// TIA Portal project "S7-1200-Single-Pump-Station" (V17)

(* hardware
DEVICE "S7-1200 station_1"  S7-1200 Station
   slot 0: "Rack_0"  S7-1200 Rack  Rack  V1.0
   slot 1: "PLC_1"  CPU 1212C DC/DC/DC  6ES7 212-1AE40-0XB0  V4.2
DEVICE "HMI_1"  TP700 Comfort
   slot 0: "HMI_1"  TP700 Comfort  6AV2 124-0GC01-0AX0  17.0.0.0
   slot 1: "HMI_RT_1"  TP700 Comfort  6AV2 124-0GC01-0AX0  17.0.0.0
   slot 5: "HMI_1.IE_CP_1"  PROFINET Interface  17.0.0.0
      slot 1: "PROFINET Interface_1"  PROFINET Interface
         slot 1: "Port_1"  Port
         slot 2: "Port_2"  Port
   slot 7: "HMI_1.MPI/DP_CP_1"  MPI/DP Interface  17.0.0.0
*)

// ===== PLC "PLC_1"  CPU 1212C DC/DC/DC =====

VAR_GLOBAL   // PLC tag table "Default tag table"
   "Clock_Byte" AT %MB100 : Byte;
   "Clock_10Hz" AT %M100.0 : Bool;
   "Clock_5Hz" AT %M100.1 : Bool;
   "Clock_2.5Hz" AT %M100.2 : Bool;
   "Clock_2Hz" AT %M100.3 : Bool;
   "Clock_1.25Hz" AT %M100.4 : Bool;
   "Clock_1Hz" AT %M100.5 : Bool;
   "Clock_0.625Hz" AT %M100.6 : Bool;
   "Clock_0.5Hz" AT %M100.7 : Bool;
   "AL" AT %I0.5 : Bool;
   "LSL" AT %I0.3 : Bool;
   "LSH" AT %I0.4 : Bool;
   "S1Auto" AT %I0.0 : Bool;
   "S2" AT %I0.2 : Bool;
   "LT" AT %IW64 : Int;
   "L1" AT %Q0.0 : Bool;
   "L2" AT %Q0.1 : Bool;
   "P1" AT %Q0.2 : Bool;
   "S1Hand" AT %I0.1 : Bool;
END_VAR

DATA_BLOCK "Random Generator DB"   // DB1
{ S7_Optimized_Access := 'TRUE' }
VERSION : 0.1
// stored: InstanceOfName Random Inflow Generator
"Random Inflow Generator"
BEGIN
END_DATA_BLOCK

DATA_BLOCK "Well DB"   // DB3
{ S7_Optimized_Access := 'TRUE' }
VERSION : 0.1
// stored: InstanceOfName Well Simulation
"Well Simulation"
BEGIN
END_DATA_BLOCK

DATA_BLOCK "Main DB"   // DB4
{ S7_Optimized_Access := 'TRUE' }
VERSION : 0.1
   VAR
      RandomInflow : Real;
      ActualInflow : Real;
      ActualOutflow : Real;
      S1AutoHMI : Bool;
      S1HandHMI : Bool;
      S2HMI : Bool;
      AutoMode : Bool;
      HandMode : Bool;
      ServiceMode : Bool;
      LevelPercent : Real;
      HighLevelReached : Bool;
      AutoPumpLatch : Bool;
      LSHHMI : Bool;
      LSLHMI : Bool;
      AlarmMode : Bool;
      HighLevelSetpoint : Real := 50.0;
      LowLevelSetpoint : Real := 20.0;
      ResetSetpoints : Bool;
      AlarmHelp : Bool := false;
      LTMeters : Real;
      ALHMI : Bool;
      PumpFault : Bool;
      HMIAlarmWord : Word;
      HighSetpointPrevious : Real := 50.0;
      LowSetpointPrevious : Real := 20.0;
      LTNormalized : Real;
      LTAnalogPercent : Real;
      SimulationMode : Bool;
      PumpStartRequest : Bool;
      PumpSafety : Bool;
      LevelInLiters : Real;
   END_VAR
BEGIN
END_DATA_BLOCK

// folder: System blocks/Program resources

DATA_BLOCK "IEC_Timer_0_DB"   // DB2
{ S7_Optimized_Access := 'TRUE' }
AUTHOR : Simatic
FAMILY : IEC
NAME : IEC_TMR
VERSION : 1.0
// stored: InstanceOfName IEC_TIMER
"IEC_TIMER"
BEGIN
END_DATA_BLOCK

DATA_BLOCK "IEC_Timer_0_DB_2"   // DB6
{ S7_Optimized_Access := 'TRUE' }
AUTHOR : Simatic
FAMILY : IEC
NAME : IEC_TMR
VERSION : 1.0
// stored: InstanceOfName IEC_TIMER
"IEC_TIMER"
BEGIN
END_DATA_BLOCK

// folder: (top level)

FUNCTION_BLOCK "Random Inflow Generator"   // FB1, LAD
{ S7_Optimized_Access := 'TRUE' }
VERSION : 0.1
   VAR_OUTPUT
      RandomInflow : Real;
   END_VAR
   VAR
      TimeStatus : Int;
      SystemTime : DTL;
      RandomValue : Int;
   END_VAR
BEGIN

REGION Network 1: System Time Acquisition
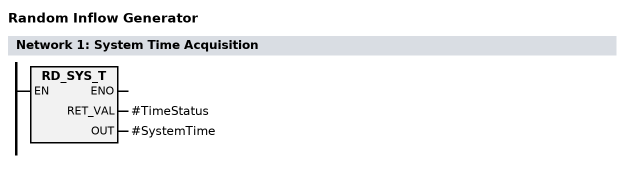
   #TimeStatus := RD_SYS_T(OUT => #SystemTime);
END_REGION

REGION Network 2 (SCL): Random Value Generation
   IF #TimeStatus = 0 THEN
       #RandomValue :=
       UDINT_TO_INT(
                     #SystemTime.NANOSECOND MOD UDINT#3
       ) + 1;
   END_IF;
END_REGION

REGION Network 3 (SCL): Random Inflow Rate Selection
   IF #RandomValue = 1 THEN
       #RandomInflow := 10.0;
   ELSIF #RandomValue = 2 THEN
       #RandomInflow := 15.0;
   ELSE
       #RandomInflow := 7.0;
   END_IF;
END_REGION
END_FUNCTION_BLOCK

FUNCTION_BLOCK "Well Simulation"   // FB2, SCL
{ S7_Optimized_Access := 'TRUE' }
VERSION : 0.1
   VAR_INPUT
      CycleTime : Real := 0.1;
      Inflow : Real;
      Outflow : Real;
   END_VAR
   VAR
      TankLevel : Real;
      ActualInflow : Real;
      ActualOutflow : Real;
      "TankLevel%" : Real;
   END_VAR
BEGIN
   #ActualOutflow := #Outflow * #CycleTime;
   #ActualInflow := #Inflow * #CycleTime;

   #TankLevel := #TankLevel + (#ActualInflow - #ActualOutflow);

   IF #TankLevel > 1250.0 THEN
       #TankLevel := 1250.0;
   END_IF;

   IF #TankLevel < 0.0 THEN
       #TankLevel := 0.0;
   END_IF;

   #"TankLevel%" := (#TankLevel / 1250.0) * 100.0;
END_FUNCTION_BLOCK

ORGANIZATION_BLOCK "Main"   // OB1, LAD, ProgramCycle
TITLE = "Main Program Sweep (Cycle)"
{ S7_Optimized_Access := 'TRUE' }
VERSION : 0.1
   VAR_INPUT
      Initial_Call : Bool;   // Initial call of this OB
      Remanence : Bool;   // =True, if remanent data are available
   END_VAR
BEGIN

REGION Network 1: LT Analog Input Scaling
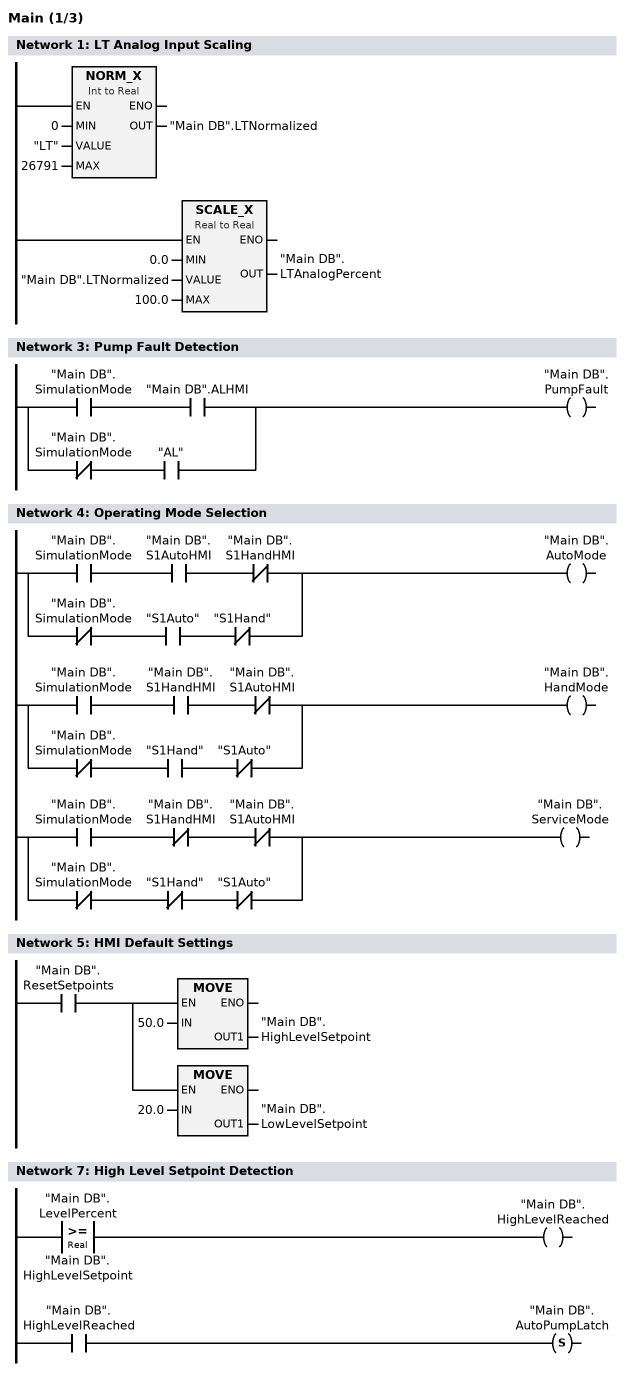
   RUNG wire#powerrail
      { S7_Templates := "[SrcType := Int, DestType := Real]" } Normalize(min := 0, value := "LT", max := 26791, out => "Main DB".LTNormalized)
   END_RUNG
   RUNG wire#powerrail
      { S7_Templates := "[SrcType := Real, DestType := Real]" } Scale(min := 0.0, value := "Main DB".LTNormalized, max := 100.0, out => "Main DB".LTAnalogPercent)
   END_RUNG
   // the same network as SCL:
   "Main DB".LTNormalized := NORM_X(MIN := 0, VALUE := "LT", MAX := 26791);
   "Main DB".LTAnalogPercent := SCALE_X(MIN := 0.0, VALUE := "Main DB".LTNormalized, MAX := 100.0);
END_REGION

REGION Network 2 (SCL): LT Source Selection and Level Conversion
   IF "Main DB".SimulationMode THEN
       "Main DB".LevelPercent := "Well DB"."TankLevel%";
       "Main DB".LevelInLiters := "Well DB".TankLevel;
   ELSE
       "Main DB".LevelPercent := "Main DB".LTAnalogPercent;
       "Main DB".LevelInLiters := ("Main DB".LevelPercent / 100.0) * 1250.0;
   END_IF;

   "Main DB".LTMeters := ("Main DB".LevelPercent * 2.5) / 100.0;
END_REGION

REGION Network 3: Pump Fault Detection
   RUNG wire#powerrail
      Contact( "Main DB".SimulationMode )
      Contact( "Main DB".ALHMI )
      wire#w1
      Coil( "Main DB".PumpFault )
   END_RUNG
   RUNG wire#powerrail
      I_Contact( "Main DB".SimulationMode )
      Contact( "AL" )
   END_RUNG wire#w1
   // the same network as SCL:
   "Main DB".PumpFault := ("Main DB".SimulationMode AND "Main DB".ALHMI) OR (NOT "Main DB".SimulationMode AND "AL");
END_REGION

REGION Network 4: Operating Mode Selection
   RUNG wire#powerrail
      Contact( "Main DB".SimulationMode )
      Contact( "Main DB".S1AutoHMI )
      I_Contact( "Main DB".S1HandHMI )
      wire#w1
      Coil( "Main DB".AutoMode )
   END_RUNG
   RUNG wire#powerrail
      I_Contact( "Main DB".SimulationMode )
      Contact( "S1Auto" )
      I_Contact( "S1Hand" )
   END_RUNG wire#w1
   RUNG wire#powerrail
      Contact( "Main DB".SimulationMode )
      Contact( "Main DB".S1HandHMI )
      I_Contact( "Main DB".S1AutoHMI )
      wire#w2
      Coil( "Main DB".HandMode )
   END_RUNG
   RUNG wire#powerrail
      I_Contact( "Main DB".SimulationMode )
      Contact( "S1Hand" )
      I_Contact( "S1Auto" )
   END_RUNG wire#w2
   RUNG wire#powerrail
      Contact( "Main DB".SimulationMode )
      I_Contact( "Main DB".S1HandHMI )
      I_Contact( "Main DB".S1AutoHMI )
      wire#w3
      Coil( "Main DB".ServiceMode )
   END_RUNG
   RUNG wire#powerrail
      I_Contact( "Main DB".SimulationMode )
      I_Contact( "S1Hand" )
      I_Contact( "S1Auto" )
   END_RUNG wire#w3
   // the same network as SCL:
   "Main DB".AutoMode := ("Main DB".SimulationMode AND "Main DB".S1AutoHMI AND NOT "Main DB".S1HandHMI) OR (NOT "Main DB".SimulationMode AND "S1Auto" AND NOT "S1Hand");
   "Main DB".HandMode := ("Main DB".SimulationMode AND "Main DB".S1HandHMI AND NOT "Main DB".S1AutoHMI) OR (NOT "Main DB".SimulationMode AND "S1Hand" AND NOT "S1Auto");
   "Main DB".ServiceMode := ("Main DB".SimulationMode AND NOT "Main DB".S1HandHMI AND NOT "Main DB".S1AutoHMI) OR (NOT "Main DB".SimulationMode AND NOT "S1Hand" AND NOT "S1Auto");
END_REGION

REGION Network 5: HMI Default Settings
   RUNG wire#powerrail
      Contact( "Main DB".ResetSetpoints )
      wire#w1
      Move(in := 50.0, out1 => "Main DB".HighLevelSetpoint)
   END_RUNG
   RUNG wire#w1
      Move(in := 20.0, out1 => "Main DB".LowLevelSetpoint)
   END_RUNG
   // the same network as SCL:
   IF "Main DB".ResetSetpoints THEN
       "Main DB".HighLevelSetpoint := 50.0;
       "Main DB".LowLevelSetpoint := 20.0;
   END_IF;
END_REGION

REGION Network 6 (SCL): HMI Setpoint Validation

   IF "Main DB".LowLevelSetpoint <> "Main DB".LowSetpointPrevious THEN

       "Main DB".LowLevelSetpoint := LIMIT(
                                           MN := 0.0,
                                           IN := "Main DB".LowLevelSetpoint,
                                           MX := "Main DB".HighLevelSetpoint - 5.0
       );

   ELSIF "Main DB".HighLevelSetpoint <> "Main DB".HighSetpointPrevious THEN

       "Main DB".HighLevelSetpoint := LIMIT(
                                            MN := "Main DB".LowLevelSetpoint + 5.0,
                                            IN := "Main DB".HighLevelSetpoint,
                                            MX := 100.0
       );

   END_IF;

   "Main DB".HighSetpointPrevious := "Main DB".HighLevelSetpoint;
   "Main DB".LowSetpointPrevious := "Main DB".LowLevelSetpoint;
END_REGION

REGION Network 7: High Level Setpoint Detection
   RUNG wire#powerrail
      { S7_Templates := "SrcType := Real" } GE_Contact(in1 := "Main DB".LevelPercent, in2 := "Main DB".HighLevelSetpoint)
      Coil( "Main DB".HighLevelReached )
   END_RUNG
   RUNG wire#powerrail
      Contact( "Main DB".HighLevelReached )
      S_Coil( "Main DB".AutoPumpLatch )
   END_RUNG
   // the same network as SCL:
   "Main DB".HighLevelReached := "Main DB".LevelPercent >= "Main DB".HighLevelSetpoint;
   IF "Main DB".HighLevelReached THEN "Main DB".AutoPumpLatch := TRUE; END_IF;
END_REGION

REGION Network 8: Low Level Setpoint Reset
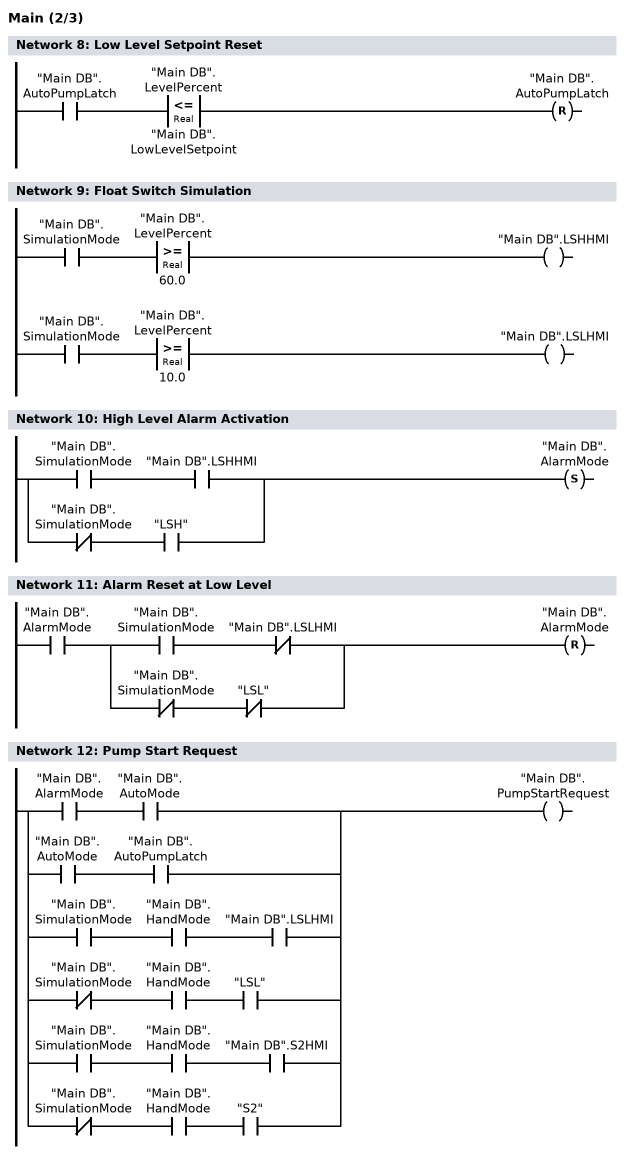
   RUNG wire#powerrail
      Contact( "Main DB".AutoPumpLatch )
      { S7_Templates := "SrcType := Real" } LE_Contact(in1 := "Main DB".LevelPercent, in2 := "Main DB".LowLevelSetpoint)
      R_Coil( "Main DB".AutoPumpLatch )
   END_RUNG
   // the same network as SCL:
   IF "Main DB".AutoPumpLatch AND ("Main DB".LevelPercent <= "Main DB".LowLevelSetpoint) THEN
       "Main DB".AutoPumpLatch := FALSE;
   END_IF;
END_REGION

REGION Network 9: Float Switch Simulation
   RUNG wire#powerrail
      Contact( "Main DB".SimulationMode )
      { S7_Templates := "SrcType := Real" } GE_Contact(in1 := "Main DB".LevelPercent, in2 := 60.0)
      Coil( "Main DB".LSHHMI )
   END_RUNG
   RUNG wire#powerrail
      Contact( "Main DB".SimulationMode )
      { S7_Templates := "SrcType := Real" } GE_Contact(in1 := "Main DB".LevelPercent, in2 := 10.0)
      Coil( "Main DB".LSLHMI )
   END_RUNG
   // the same network as SCL:
   "Main DB".LSHHMI := "Main DB".SimulationMode AND ("Main DB".LevelPercent >= 60.0);
   "Main DB".LSLHMI := "Main DB".SimulationMode AND ("Main DB".LevelPercent >= 10.0);
END_REGION

REGION Network 10: High Level Alarm Activation
   RUNG wire#powerrail
      Contact( "Main DB".SimulationMode )
      Contact( "Main DB".LSHHMI )
      wire#w1
      S_Coil( "Main DB".AlarmMode )
   END_RUNG
   RUNG wire#powerrail
      I_Contact( "Main DB".SimulationMode )
      Contact( "LSH" )
   END_RUNG wire#w1
   // the same network as SCL:
   IF ("Main DB".SimulationMode AND "Main DB".LSHHMI) OR (NOT "Main DB".SimulationMode AND "LSH") THEN
       "Main DB".AlarmMode := TRUE;
   END_IF;
END_REGION

REGION Network 11: Alarm Reset at Low Level
   RUNG wire#powerrail
      Contact( "Main DB".AlarmMode )
      wire#w1
      Contact( "Main DB".SimulationMode )
      I_Contact( "Main DB".LSLHMI )
      wire#w2
      R_Coil( "Main DB".AlarmMode )
   END_RUNG
   RUNG wire#w1
      I_Contact( "Main DB".SimulationMode )
      I_Contact( "LSL" )
   END_RUNG wire#w2
   // the same network as SCL:
   IF "Main DB".AlarmMode AND (("Main DB".SimulationMode AND NOT "Main DB".LSLHMI) OR (NOT "Main DB".SimulationMode AND NOT "LSL")) THEN
       "Main DB".AlarmMode := FALSE;
   END_IF;
END_REGION

REGION Network 12: Pump Start Request
   RUNG wire#powerrail
      Contact( "Main DB".AlarmMode )
      Contact( "Main DB".AutoMode )
      wire#w1
      Coil( "Main DB".PumpStartRequest )
   END_RUNG
   RUNG wire#powerrail
      Contact( "Main DB".AutoMode )
      Contact( "Main DB".AutoPumpLatch )
   END_RUNG wire#w1
   RUNG wire#powerrail
      Contact( "Main DB".SimulationMode )
      Contact( "Main DB".HandMode )
      Contact( "Main DB".LSLHMI )
   END_RUNG wire#w1
   RUNG wire#powerrail
      I_Contact( "Main DB".SimulationMode )
      Contact( "Main DB".HandMode )
      Contact( "LSL" )
   END_RUNG wire#w1
   RUNG wire#powerrail
      Contact( "Main DB".SimulationMode )
      Contact( "Main DB".HandMode )
      Contact( "Main DB".S2HMI )
   END_RUNG wire#w1
   RUNG wire#powerrail
      I_Contact( "Main DB".SimulationMode )
      Contact( "Main DB".HandMode )
      Contact( "S2" )
   END_RUNG wire#w1
   // the same network as SCL:
   "Main DB".PumpStartRequest := ("Main DB".AlarmMode AND "Main DB".AutoMode) OR ("Main DB".AutoMode AND "Main DB".AutoPumpLatch) OR ("Main DB".SimulationMode AND "Main DB".HandMode AND "Main DB".LSLHMI) OR (NOT "Main DB".SimulationMode AND "Main DB".HandMode AND "LSL") OR ("Main DB".SimulationMode AND "Main DB".HandMode AND "Main DB".S2HMI) OR (NOT "Main DB".SimulationMode AND "Main DB".HandMode AND "S2");
END_REGION

REGION Network 13: Pump Safety Interlocks
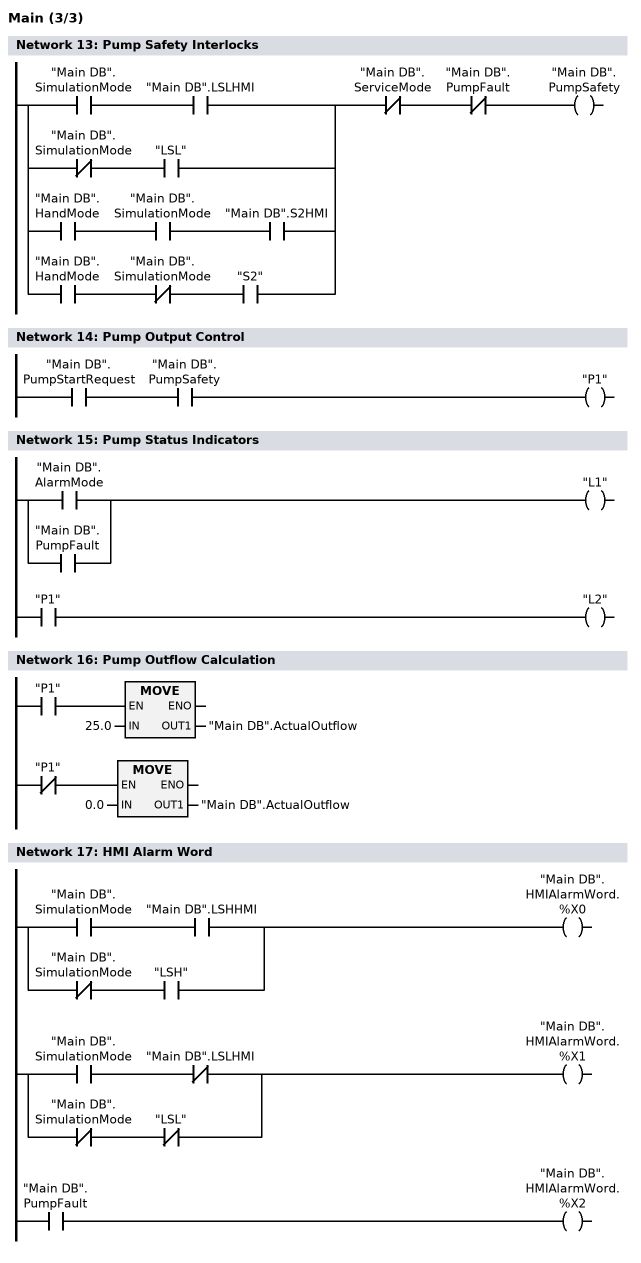
   RUNG wire#powerrail
      Contact( "Main DB".SimulationMode )
      Contact( "Main DB".LSLHMI )
      wire#w1
      I_Contact( "Main DB".ServiceMode )
      I_Contact( "Main DB".PumpFault )
      Coil( "Main DB".PumpSafety )
   END_RUNG
   RUNG wire#powerrail
      I_Contact( "Main DB".SimulationMode )
      Contact( "LSL" )
   END_RUNG wire#w1
   RUNG wire#powerrail
      Contact( "Main DB".HandMode )
      Contact( "Main DB".SimulationMode )
      Contact( "Main DB".S2HMI )
   END_RUNG wire#w1
   RUNG wire#powerrail
      Contact( "Main DB".HandMode )
      I_Contact( "Main DB".SimulationMode )
      Contact( "S2" )
   END_RUNG wire#w1
   // the same network as SCL:
   "Main DB".PumpSafety := (("Main DB".SimulationMode AND "Main DB".LSLHMI) OR (NOT "Main DB".SimulationMode AND "LSL") OR ("Main DB".HandMode AND "Main DB".SimulationMode AND "Main DB".S2HMI) OR ("Main DB".HandMode AND NOT "Main DB".SimulationMode AND "S2")) AND NOT "Main DB".ServiceMode AND NOT "Main DB".PumpFault;
END_REGION

REGION Network 14: Pump Output Control
   RUNG wire#powerrail
      Contact( "Main DB".PumpStartRequest )
      Contact( "Main DB".PumpSafety )
      Coil( "P1" )
   END_RUNG
   // the same network as SCL:
   "P1" := "Main DB".PumpStartRequest AND "Main DB".PumpSafety;
END_REGION

REGION Network 15: Pump Status Indicators
   RUNG wire#powerrail
      Contact( "Main DB".AlarmMode )
      wire#w1
      Coil( "L1" )
   END_RUNG
   RUNG wire#powerrail
      Contact( "Main DB".PumpFault )
   END_RUNG wire#w1
   RUNG wire#powerrail
      Contact( "P1" )
      Coil( "L2" )
   END_RUNG
   // the same network as SCL:
   "L1" := "Main DB".AlarmMode OR "Main DB".PumpFault;
   "L2" := "P1";
END_REGION

REGION Network 16: Pump Outflow Calculation
   RUNG wire#powerrail
      Contact( "P1" )
      Move(in := 25.0, out1 => "Main DB".ActualOutflow)
   END_RUNG
   RUNG wire#powerrail
      I_Contact( "P1" )
      Move(in := 0.0, out1 => "Main DB".ActualOutflow)
   END_RUNG
   // the same network as SCL:
   IF "P1" THEN "Main DB".ActualOutflow := 25.0; END_IF;
   IF NOT "P1" THEN "Main DB".ActualOutflow := 0.0; END_IF;
END_REGION

REGION Network 17: HMI Alarm Word
   RUNG wire#powerrail
      Contact( "Main DB".SimulationMode )
      Contact( "Main DB".LSHHMI )
      wire#w1
      Coil( "Main DB".HMIAlarmWord.%X0 )
   END_RUNG
   RUNG wire#powerrail
      I_Contact( "Main DB".SimulationMode )
      Contact( "LSH" )
   END_RUNG wire#w1
   RUNG wire#powerrail
      Contact( "Main DB".SimulationMode )
      I_Contact( "Main DB".LSLHMI )
      wire#w2
      Coil( "Main DB".HMIAlarmWord.%X1 )
   END_RUNG
   RUNG wire#powerrail
      I_Contact( "Main DB".SimulationMode )
      I_Contact( "LSL" )
   END_RUNG wire#w2
   RUNG wire#powerrail
      Contact( "Main DB".PumpFault )
      Coil( "Main DB".HMIAlarmWord.%X2 )
   END_RUNG
   // the same network as SCL:
   "Main DB".HMIAlarmWord.%X0 := ("Main DB".SimulationMode AND "Main DB".LSHHMI) OR (NOT "Main DB".SimulationMode AND "LSH");
   "Main DB".HMIAlarmWord.%X1 := ("Main DB".SimulationMode AND NOT "Main DB".LSLHMI) OR (NOT "Main DB".SimulationMode AND NOT "LSL");
   "Main DB".HMIAlarmWord.%X2 := "Main DB".PumpFault;
END_REGION
END_ORGANIZATION_BLOCK

ORGANIZATION_BLOCK "Well Cycle"   // OB30, LAD, CyclicInterrupt
{ S7_Optimized_Access := 'TRUE' }
VERSION : 0.1
   VAR_INPUT
      Initial_Call : Bool;   // Initial call of this OB
      Event_Count : Int;   // Events discarded
   END_VAR
BEGIN

REGION Network 1: Well Level Simulation
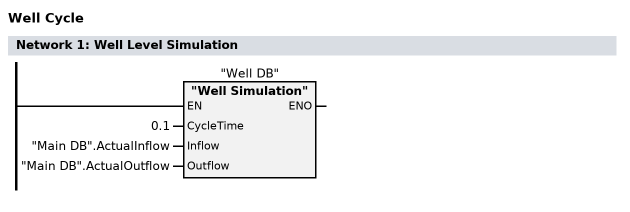
   RUNG wire#powerrail
      "Well DB"(CycleTime := 0.1, Inflow := "Main DB".ActualInflow, Outflow := "Main DB".ActualOutflow)
   END_RUNG
   // the same network as SCL:
   "Well DB"(CycleTime := 0.1, Inflow := "Main DB".ActualInflow, Outflow := "Main DB".ActualOutflow);   // "Well Simulation"
END_REGION
END_ORGANIZATION_BLOCK

ORGANIZATION_BLOCK "Inflow Generator"   // OB123, LAD, ProgramCycle
TITLE = "Main Program Sweep (Cycle)"
{ S7_Optimized_Access := 'TRUE' }
VERSION : 0.1
   VAR_INPUT
      Initial_Call : Bool;   // Initial call of this OB
      Remanence : Bool;   // =True, if remanent data are available
   END_VAR
BEGIN

REGION Network 1: Random Inflow Generator Call
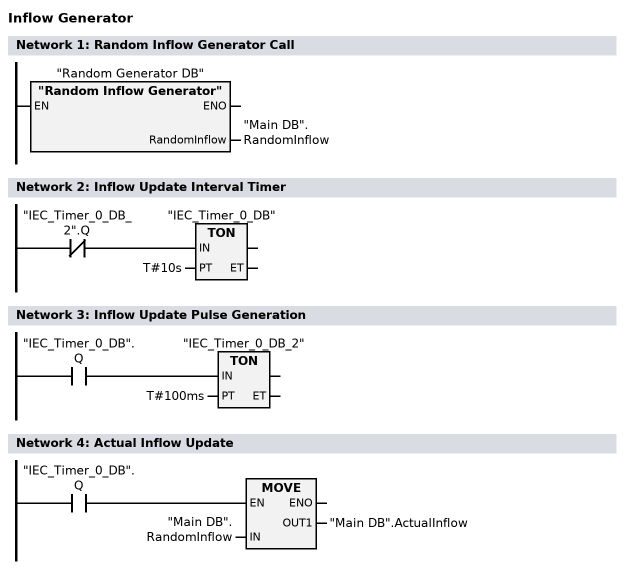
   RUNG wire#powerrail
      "Random Generator DB"(RandomInflow => "Main DB".RandomInflow)
   END_RUNG
   // the same network as SCL:
   "Random Generator DB"(RandomInflow => "Main DB".RandomInflow);   // "Random Inflow Generator"
END_REGION

REGION Network 2: Inflow Update Interval Timer
   "IEC_Timer_0_DB".TON(IN := NOT "IEC_Timer_0_DB_2".Q, PT := T#10s);
END_REGION

REGION Network 3: Inflow Update Pulse Generation
   "IEC_Timer_0_DB_2".TON(IN := "IEC_Timer_0_DB".Q, PT := T#100ms);
END_REGION

REGION Network 4: Actual Inflow Update
   RUNG wire#powerrail
      Contact( "IEC_Timer_0_DB".Q )
      Move(in := "Main DB".RandomInflow, out1 => "Main DB".ActualInflow)
   END_RUNG
   // the same network as SCL:
   IF "IEC_Timer_0_DB".Q THEN "Main DB".ActualInflow := "Main DB".RandomInflow; END_IF;
END_REGION
END_ORGANIZATION_BLOCK

(* ===== HMI "HMI_RT_1" =====
system functions are stored by id; their names below are inferred from use
connection "HMI_Connection_1": ETHERNET, S7_1200_OMS

HMI tags "Default tag table"
   "Tag_ScreenNumber" : UInt, internal
   "Well DB_TankLevel" : Real = PLC "Well DB".TankLevel, 1 s
   "Main DB_AutoMode" : Bool = PLC "Main DB".AutoMode, 1 s
   "Main DB_HandMode" : Bool = PLC "Main DB".HandMode, 1 s
   "Main DB_S1Auto" : Bool = PLC "Main DB".S1AutoHMI, 1 s
   "Main DB_S1Hand" : Bool = PLC "Main DB".S1HandHMI, 1 s
   "Main DB_MaintainMode" : Bool = PLC "Main DB".ServiceMode, 1 s
   "Main DB_S2" : Bool = PLC "Main DB".S2HMI, 1 s
   "Liters/%" : Bool AT %DB1.DBX0.0
   "Well DB_TankLevel%" : Real = PLC "Well DB".TankLevel%, 1 s
   "Well DB_ActualInflow" : Real = PLC "Well DB".ActualInflow, 1 s
   "Well DB_ActualOutflow" : Real = PLC "Well DB".ActualOutflow, 1 s
   "Main DB_LT" : Real = PLC "Main DB".LevelPercent, 1 s
   "Well DB_Inflow" : Real = PLC "Well DB".Inflow, 1 s
   "Well DB_Outflow" : Real = PLC "Well DB".Outflow, 1 s
   "Main DB_LT_HMI_H" : Real = PLC "Main DB".HighLevelSetpoint, 1 s
   "Main DB_LT_HMI_L" : Real = PLC "Main DB".LowLevelSetpoint, 1 s
   "Main DB_ResetSetpoints" : Bool = PLC "Main DB".ResetSetpoints, 1 s
   "ResetSetpoints" : Bool AT %DB1.DBX0.0
   "Main DB_LSH" : Bool = PLC "Main DB".LSHHMI, 1 s
   "Main DB_LSL" : Bool = PLC "Main DB".LSLHMI, 1 s
   "Main DB_AlarmHelp" : Bool = PLC "Main DB".AlarmHelp, 1 s
   "Main DB_AlarmMode" : Bool = PLC "Main DB".AlarmMode, 1 s
   "Main DB_LT_Meters" : Real = PLC "Main DB".LTMeters, 1 s
   "Meters/%" : Bool AT %DB1.DBX0.0
   "Main DB_PumpFault" : Bool = PLC "Main DB".PumpFault, 1 s
   "Main DB_HMI_AlarmWord" : Word = PLC "Main DB".HMIAlarmWord, 1 s
   "Main DB_AL" : Bool = PLC "Main DB".ALHMI, 1 s
   "L1" : Bool = PLC L1 AT %Q0.0, 1 s
   "L2" : Bool = PLC L2 AT %Q0.1, 1 s
   "Main DB_SimulationMode" : Bool = PLC "Main DB".SimulationMode, 1 s
   "Main DB_LevelInLiters" : Real = PLC "Main DB".LevelInLiters, 1 s

discrete alarms
   1: 'High water level', class Errors, trigger "Main DB_HMI_AlarmWord" bit 0
   2: 'Low water level', class Warnings, trigger "Main DB_HMI_AlarmWord" bit 1
   3: 'Pump stopped', class Errors, trigger "Main DB_HMI_AlarmWord" bit 2

screen "Tank Control" 800x420, template "Template_1"
   on GenerateScreen: SetTag("Tag_ScreenNumber", 1)
   Bar "Bar_1" at 319,68 size 157x267; MinimumValue 0; MaximumValue 1250
      Visibility <- "Liters/%"
      ProcessValue <- "Main DB_LevelInLiters"
   Circle "Circle_1" at 111,143 size 48x48
      Appearance <- "Main DB_MaintainMode"
   Button "Button_3" at 11,152 size 96x32; TextOff 'Service'
      on Click: ResetBit("Main DB_S1Auto"); ResetBit("Main DB_S1Hand")
      ObjectEnable <- "Main DB_SimulationMode"
   Circle "Circle_2" at 111,93 size 48x48
      Visibility <- "Main DB_HandMode"
   Button "Button_1" at 11,102 size 96x32; TextOff 'Hand'
      on Click: SetBit("Main DB_S1Hand"); ResetBit("Main DB_S1Auto")
      ObjectEnable <- "Main DB_SimulationMode"
   Circle "Circle_3" at 111,43 size 48x48
      Appearance <- "Main DB_AutoMode"
   Button "Button_2" at 11,52 size 96x32; TextOff 'Auto'
      on Click: SetBit("Main DB_S1Auto"); ResetBit("Main DB_S1Hand")
      ObjectEnable <- "Main DB_SimulationMode"
   Circle "Circle_5" at 214,93 size 48x48
      Visibility <- "Main DB_HandMode"
      Appearance <- "Main DB_HandMode"
   Button "Button_5" at 114,102 size 96x32; TextOff 'Pump'
      on Press: SetBit("Main DB_S2")
      on Release: ResetBit("Main DB_S2")
      Visibility <- "Main DB_HandMode"
      ObjectEnable <- "Main DB_SimulationMode"
   Switch "Switch_1" at 408,12 size 66x49; CaptionText 'Switch'; TextOff '%'; TextOn 'Liters'
      ProcessValue <- "Liters/%"
   TextField "Text field_1" at 322,17 size 76x40; Text 'Well'
   Bar "Bar_2" at 319,68 size 157x267; MinimumValue 0; MaximumValue 100
      Visibility <- "Liters/%"
      ProcessValue <- "Main DB_LT"
   IOField "I/O field_1" at 648,179 size 34x32; FormatPattern 9999999
      ProcessValue <- "Well DB_Inflow"
   TextField "Text field_2" at 589,184 size 63x23; Text 'Inflow'
   TextField "Text field_3" at 683,183 size 30x23; Text 'l/s'
   IOField "I/O field_2" at 659,219 size 34x32; FormatPattern 9999999
      ProcessValue <- "Well DB_Outflow"
   TextField "Text field_4" at 589,224 size 76x23; Text 'Outflow'
   TextField "Text field_5" at 694,224 size 30x23; Text 'l/s'
   IOField "I/O field_3" at 673,259 size 45x32; FormatPattern 999
      ProcessValue <- "Main DB_LT"
      Visibility <- "Meters/%"
   TextField "Text field_6" at 589,264 size 92x23; Text 'LT sensor'
   TextField "Text field_8" at 5,262 size 100x23; Text 'LT Level H'
   IOField "I/O field_4" at 101,257 size 35x32; FormatPattern 99
      ProcessValue <- "Main DB_LT_HMI_H"
   TextField "Text field_9" at 5,313 size 97x23; Text 'LT Level L'
   IOField "I/O field_5" at 101,308 size 35x32; FormatPattern 99
      ProcessValue <- "Main DB_LT_HMI_L"
   Button "Button_4" at 177,257 size 135x85; TextOff 'Default settings'
      on Press: SetBit("Main DB_ResetSetpoints"); SetBit("ResetSetpoints"); SetBit("Main DB_S1Auto"); ResetBit("Main DB_S1Hand"); ResetBit("Main DB_PumpFault")
      on Release: ResetBit("Main DB_ResetSetpoints")
      Visibility <- "ResetSetpoints"
   TextField "Text field_10" at 589,298 size 39x23; Text 'LSH'
   Circle "Circle_4" at 627,295 size 28x28
      Appearance <- "Main DB_HMI_AlarmWord"
   TextField "Text field_11" at 589,335 size 36x23; Text 'LSL'
   Circle "Circle_6" at 627,332 size 28x28
      Appearance <- "Main DB_HMI_AlarmWord"
   Circle "Circle_7" at 111,193 size 48x48
      Appearance <- "Main DB_AlarmMode"
   Button "Button_6" at 11,202 size 96x32; TextOff 'Alarm'
      ObjectEnable <- "Main DB_AlarmHelp"
   TextField "Text field_12" at 589,84 size 55x23; Text 'Pump'
   Circle "Circle_8" at 640,70 size 48x48
      Appearance <- "L2"
   Switch "Switch_2" at 723,259 size 34x32; CaptionText 'Switch'; TextOff '%'; TextOn 'm'
      ProcessValue <- "Meters/%"
   IOField "I/O field_6" at 673,259 size 49x32; FormatPattern 9.99
      ProcessValue <- "Main DB_LT_Meters"
      Visibility <- "Meters/%"
   TextField "Text field_7" at 588,134 size 104x23; Text 'Pump fault'
   Circle "Circle_9" at 683,120 size 48x48
      Appearance <- "Main DB_PumpFault"
   TextField "Text field_13" at 17,12 size 84x34; Text 'MODE'
   TextField "Text field_14" at 589,34 size 59x23; Text 'Alarm'
   Circle "Circle_10" at 648,21 size 48x48
      Appearance <- "L1"
   Switch "Switch_3" at 734,126 size 37x39; CaptionText 'Switch'; TextOff 'OFF'; TextOn 'ON'
      ProcessValue <- "Main DB_AL"
      ObjectEnable <- "Main DB_SimulationMode"
   TextField "Text field_15" at 136,262 size 25x23; Text '%'
   TextField "Text field_16" at 134,313 size 25x23; Text '%'
   TextField "Text field_17" at 195,230 size 102x23; Text 'Simulation'
      Visibility <- "ResetSetpoints"
   Switch "Switch_4" at 177,257 size 135x85; CaptionText 'Switch'; TextOff 'OFF'; TextOn 'ON'
      ProcessValue <- "Main DB_SimulationMode"
      Visibility <- "ResetSetpoints"

Template "Template_1" 800x420
   Button "Exit" at 720,360 size 78x58; TextOff 'Exit'; PictureOff "ExitRuntime_TP700_Comfort_TR"; PictureOn "ExitRuntime_TP700_Comfort_TR"
      on Release: StopRuntime(0)
   Button "Template_Button_7" at 81,360 size 78x58; TextOff 'Alarms'
      on Release: ActivateScreen("Alarms", 1)
   Button "Start screen" at 1,360 size 78x58; TextOff 'Start screen'; PictureOff "NavigateHome_TP700_Comfort_TR"; PictureOn "NavigateHome_TP700_Comfort_TR"
      on Release: ActivateScreen("Tank Control", 0)

screen "Alarms" 800x420, template "Template_1"
   AlarmView "Alarm view_1" at 3,1 size 793x357
*)